PROGRAM P_BeamClassAssertion
VAR
    {attribute 'pytmc' := '
    pv: @(PREFIX)BeamClassWatcher
    '}
    fbBeamClassWatcher : FB_BeamClassWatcher;
    {attribute 'pytmc' := '
    pv: @(PREFIX)BeamClassOutputs
    '}
    fbMPSInterface	:	FB_BeamClassOutputs_BCD;

END_VAR


// Request beam class
fbMPSInterface(BP := PMPS_GVL.stRequestedBeamParameters);

// Keep an eye on the beam class
fbBeamClassWatcher(i_stCurrentBeamParams	:= PMPS_GVL.stCurrentBeamParameters,
                    i_stRequestedBeamParams := PMPS_GVL.stRequestedBeamParameters,
                    io_fbFFHWO:= GVL.g_FastFaultOutput1,
                    i_xAutoReset := TRUE);

END_PROGRAM

(* stored: Version 1.1.0.1, ProductVersion 3.1.4022.18
   POU P_BeamClassAssertion: Id {60648296-2385-4133-a8e3-f7d1443b93ab}, SpecialFunc None *)
